(* IEC 61131-3 sources: rusty/tests/lit/multi/parse_errors_reported_once, 2 files *)

(* ---- first.st ---- *)
FUNCTION first : BOOL
VAR_INPUT
    in : BOOL;
    in2
END_VAR
;
END_FUNCTION

(* ---- second.st ---- *)
FUNCTION second : DINT
    second := 2 *;
END_FUNCTION
